// Événement d'alarme du tampon circulaire (docs/14 § 5)
{attribute 'pack_mode' := '1'}
TYPE ST_AlarmEventRec :
STRUCT
    nSeq : UDINT;
    eEvent : E_AlarmEvent;
    tTime : LINT;
    stAlarm : ST_AlarmEntry;
    sUser : STRING(24);
END_STRUCT
END_TYPE

(* stored: Version 1.1.0.1, ProductVersion 3.1.4024.12
   DUT ST_AlarmEventRec: Id {d2adea1c-4c85-5f3a-8699-e7fb8486ca37} *)
